Fanuc KAREL source: kf00105.KL

-- PROVISIONAL review KL for V770-1; original PC SHA256 cee6b260c7986a33a9efedb36e0dfbfdd90ebc4ce31aeb157af1a36b031d43c7
-- Incomplete behavior may be omitted. Consult companion uncertainty JSON. Do not deploy.
PROGRAM KF00105
%NOLOCKGROUP
BEGIN
  -- UNRESOLVED_PC offsets 5-16; opcodes 2E,23
  -- UNRESOLVED_PC offsets 21-32; opcodes 2E,23
  -- UNRESOLVED_PC offsets 37-57; opcodes 27,27,9D,22,2A,22,31
  -- UNRESOLVED_PC offsets 62-66; opcodes 7F
END KF00105
